Fanuc KAREL source: KT00982.KL

PROGRAM KT00982
%NOLOCKGROUP
VAR
  R1: REAL
  R2: REAL
  CFG: CONFIG
  OUT: POSITION
BEGIN
  R1 = 2.0
  R2 = 3.0
  R1 = 2.0
  R2 = 3.0
  CFG.CFG_FLIP = TRUE
  OUT = POS(R1, R1, R1, R1, R1, R1, CFG)
END KT00982
